TYPE ST_EL2904_A :
STRUCT
    sTerminalName       	: STRING(80) := 'EL2904 | 4-Channel Safety Digital Output';
    
    // TwinSAFE physical hardware channels (Safe Outputs 1 to 4)
    qEL2904_Ch1 				AT %Q*	: 	BOOL;	// EL2904 channel 1
	qEL2904_Ch2					AT %Q* 	: 	BOOL;	// EL2904 channel 2
	qEL2904_Ch3             	AT %Q*	: 	BOOL;	// EL2904 channel 3 			
	qEL2904_Ch4      			AT %Q*  : 	BOOL;	// EL2904 channel 4 
    
    // Hardware status and diagnostic signals
    bError              	: BOOL; // TRUE if a fault is detected (short-circuit, overload, or FSoE error)
    bReady              	: BOOL; // TRUE if terminal is active and TwinSAFE communication is OK
	
	stTerminalInfo			: 	ST_Terminal_Info;
END_STRUCT
END_TYPE

(* stored: Version 1.1.0.1
   DUT ST_EL2904_A: Id {b47fa1ee-8218-430d-bdaf-20385f9eef63} *)
